(* IEC 61131-3 sources: kns-port-domestic/tools/plcopen/tests/fixtures/constructs/src/DUTs/Motor, 1 file *)

(* ---- ST_MotorCmd.dut.st ---- *)
// Команды двигателя от HMI (DUT в папке проекта)
TYPE ST_MotorCmd :
STRUCT
    xStart : BOOL;
    xStop : BOOL;
    eMode : E_Mode := E_Mode.OutOfService;
END_STRUCT
END_TYPE
